FUNCTION_BLOCK INIT_ON_OFF (* E_TRIG Counterpart, erweitert um zwei eigenstaendige Pass-Throughs INIT_ON/INITO_ON (EInitOn) und INIT_OFF/INITO_OFF (EInitOff) *)
  (* Standard: 61131-3; Classification: standard boolean function; Description: Copyright (c) 2026 Meisterschulen am Ostbahnhof This program and the accompanying materials are made available under the terms of the Eclipse Public License 2.0 which is available at https://www.eclipse.org/legal/epl-2.0/ SPDX-License-Identifier: EPL-2.0 *)
  (* Version 1.0, 2026-10-11, Franz Höpfinger, Meisterschulen am Ostbahnhof, initial API and implementation and/or initial documentation. Basiert auf dem INIT.fbt Pass-Through-Muster, vereint die beiden Zusatzkanaele aus INIT_ON.fbt und INIT_OFF.fbt in einem FB. *)
  PACKAGE events::init;
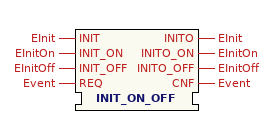
  EVENT_INPUT
    INIT : EInit; (* Initialization Request *)
    INIT_ON : EInitOn; (* Initialization Request, eigener Kanal unabhaengig von INIT *)
    INIT_OFF : EInitOff; (* Initialization Request, eigener Kanal unabhaengig von INIT *)
    REQ; (* Service Request *)
  END_EVENT
  EVENT_OUTPUT
    INITO : EInit; (* Initialization Confirm *)
    INITO_ON : EInitOn; (* Initialization Confirm, eigener Kanal unabhaengig von INITO *)
    INITO_OFF : EInitOff; (* Initialization Confirm, eigener Kanal unabhaengig von INITO *)
    CNF; (* Confirmation of Requested Service *)
  END_EVENT
  EVENT_CONNECTIONS
    INIT TO INITO;
    REQ TO CNF;
    INIT_ON TO INITO_ON;
    INIT_OFF TO INITO_OFF;
  END_CONNECTIONS
END_FUNCTION_BLOCK
